TYPE ST_STOEBERSI6SC6CIA402_REF : FB_STOEBERSI6SC6CIA402_REF;
END_TYPE

(* stored: Version 1.1.0.1, ProductVersion 3.1.4024.15
   DUT ST_STOEBERSI6SC6CIA402_REF: Id {aec84d97-c686-4afa-9bd6-0a1918754958} *)
